// TIA Portal V21 export
FUNCTION_BLOCK "FB_SclTimers"   // FB2, SCL
TITLE = IEC timers, counters and edges
{ S7_Optimized_Access := 'TRUE' }
// Every IEC timer, edge and counter as a multi-instance, each called every cycle
// stored: MemoryReserve 100, SetENOAutomatically false
   VAR_INPUT
      Start : Bool;   // Start signal
      Reset : Bool;   // Reset the counter
      DelayTime : Time := T#2S;   // On-delay time
   END_VAR
   VAR_OUTPUT
      DelayedOn : Bool;   // Start delayed by DelayTime
      RunOn : Bool;   // Start with run-on time
      Pulse : Bool;   // Pulse on the rising edge of Start
      Count : Int;   // Number of falling edges of Start
      CountReached : Bool;   // Count has reached the preset
   END_VAR
   VAR
      OnDelay { S7_SetPoint := 'True'} : TON_TIME;   // On-delay timer
      OffDelay { S7_SetPoint := 'True'} : TOF_TIME;   // Off-delay timer
      PulseTimer { S7_SetPoint := 'True'} : TP_TIME;   // Pulse timer
      StartEdge { S7_SetPoint := 'True'} : R_TRIG;   // Rising edge of Start
      StopEdge { S7_SetPoint := 'True'} : F_TRIG;   // Falling edge of Start
      PartCounter { S7_SetPoint := 'True'} : CTU_INT;   // Up counter
   END_VAR
   VAR CONSTANT
      COUNT_PRESET : Int := 10;   // Counter preset
   END_VAR
BEGIN

       REGION Timers
           #OnDelay(IN := #Start, PT := #DelayTime, Q => #DelayedOn);
           #OffDelay(IN := #Start, PT := T#3s, Q => #RunOn);
       END_REGION

       REGION Edges and pulse
           #StartEdge(CLK := #Start);
           #StopEdge(CLK := #Start);
           #PulseTimer(IN := #StartEdge.Q, PT := T#500ms, Q => #Pulse);
       END_REGION

       REGION Counter
           #PartCounter(CU := #StopEdge.Q, R := #Reset, PV := #COUNT_PRESET, Q => #CountReached, CV => #Count);
       END_REGION
END_FUNCTION_BLOCK
